Staubli VAL3: click_refreshAllMsg.pgx

program click_refreshAllMsg()
begin
  nMsgType=0
  call initMsg()
  call rs:getLog(sRobotMsg,nMsgType)
  userPageSet("message","btnAllMsg","style.backgroundColor","#33FF33")
  userPageSet("message","btnRobotMsg","style.backgroundColor","#FFFFFF")
  userPageSet("message","btnTrajMsg","style.backgroundColor","#FFFFFF")
  userPageSet("message","btnIOMsg","style.backgroundColor","#FFFFFF")
end
